Staubli VAL3: insertDelay.pgx

public program insertDelay()
  local bool l_bExit
  local bool l_bResult
  local num l_nPoint
begin
  do

    if util:sPage!="insertDelay"
      util:sPage="insertDelay"
      nSetDelay=0
      userPageBindClick("insertDelay","btn1",bConfirmDelay,true)
      userPageBindClick("insertDelay","btn2",bBackDelay,true)
      userPageBind("insertDelay","nmb1","value",nSetDelay,1,"rw")
      userPage(util:sPage)
      delay(0.5)

    endIf


    if bConfirmDelay
      bConfirmDelay=false
       call trajectory:getPointIndex(sTrajItem,sSelPoint,l_nPoint,l_bResult)
      call trajectory:insertDelay(sTrajItem,l_nPoint,bToSave,7,nSetDelay)
      l_bExit=true

    elseIf bBackDelay
      bBackDelay=false
      l_bExit=true
    endIf




    delay(0)
  until l_bExit==true
end
